Fanuc KAREL source: KT00546.KL

PROGRAM KT00546
%NOLOCKGROUP
VAR
  P1: JOINTPOS
  P2: XYZWPREXT
  OUT: XYZWPREXT
BEGIN
    P2.Y = 2.0
  OUT = P1 : P2
END KT00546
